(* PLC project g_two_hand, Anonymous Benchmark Suite 1.0 *)
(* stored: creationDateTime 2026-08-28T00:00:00 *)

PROGRAM g_two_hand
  VAR_INPUT
    LH : BOOL;
    RH : BOOL;
  END_VAR
  VAR_OUTPUT
    BothOff : BOOL;
    Armed : BOOL;
    Stroke : BOOL;
  END_VAR

(* LD diagram, written out as Structured Text *)
BothOff := NOT LH AND NOT RH;
Armed := (Armed OR BothOff) AND NOT Stroke;
Stroke := (Stroke OR Armed) AND LH AND RH;
END_PROGRAM

CONFIGURATION Config0
  RESOURCE Res0 ON PLC
    TASK tcyclic(INTERVAL := T#10ms, PRIORITY := 0);
    PROGRAM inst0 WITH tcyclic : g_two_hand;
  END_RESOURCE
END_CONFIGURATION
